// TIA Portal V20 export
Screen "Grinding"  395x400
  ScreenItem "Robot Name" at 2,2 size 393x48  Type=HmiIOField
  ScreenItem "Background" at -24,46 size 419x350  Type=HmiRectangle
  ScreenItem "Cancel Mode" at 315,4 size 76x42  Type=HmiButton
  ScreenItem "矩形_4" at 31,58 size 324x319  Type=HmiRectangle
  ScreenItem "Text Filed E- Stop_17" at 39,323 size 148x21  Type=HmiTextBox
  ScreenItem "Text Field In Auto On_9" at 39,88 size 148x21  Type=HmiTextBox
  ScreenItem "Text Field Home Position_17" at 39,111 size 148x21  Type=HmiTextBox
  ScreenItem "Text field Robot Status_5" at 33,59 size 324x26  Type=HmiTextBox
  ScreenItem "Text Field Manual_17" at 39,253 size 148x21  Type=HmiTextBox
  ScreenItem "Text Field System Ready_9" at 39,135 size 148x21  Type=HmiTextBox
  ScreenItem "Text Field Motor On_9" at 39,158 size 148x21  Type=HmiTextBox
  ScreenItem "Text Field In Cycle_9" at 39,182 size 148x21  Type=HmiTextBox
  ScreenItem "Text Field Cycle On_17" at 39,205 size 148x21  Type=HmiTextBox
  ScreenItem "Text Field On Path_17" at 39,229 size 148x21  Type=HmiTextBox
  ScreenItem "Text Field Tryout Mode_17" at 39,276 size 148x21  Type=HmiTextBox
  ScreenItem "Text Field Stop_17" at 39,300 size 148x21  Type=HmiTextBox
  ScreenItem "Text Filed Error_9" at 39,347 size 148x21  Type=HmiTextBox
  ScreenItem "Text Filed Process Fault_9" at 197,88 size 148x21  Type=HmiTextBox
  ScreenItem "Text Field Home Position_18" at 197,112 size 148x21  Type=HmiTextBox
  ScreenItem "Text Filed E- Stop_18" at 197,254 size 148x21  Type=HmiTextBox
  ScreenItem "Text Field Manual_18" at 197,183 size 148x21  Type=HmiTextBox
  ScreenItem "Text Field Cycle On_18" at 197,136 size 148x21  Type=HmiTextBox
  ScreenItem "Text Field On Path_18" at 197,159 size 148x21  Type=HmiTextBox
  ScreenItem "Text Field Tryout Mode_18" at 197,206 size 148x21  Type=HmiTextBox
  ScreenItem "Text Field Stop_18" at 197,230 size 148x21  Type=HmiTextBox
  ScreenItem "Text Field In Auto On_10" at 197,277 size 148x21  Type=HmiTextBox
  ScreenItem "Text Field Home Position_19" at 197,300 size 148x21  Type=HmiTextBox
  ScreenItem "Text Field System Ready_10" at 197,324 size 148x21  Type=HmiTextBox
  ScreenItem "Text Field Motor On_10" at 197,347 size 148x21  Type=HmiTextBox
